Staubli VAL3: stop.pgx

program stop()
// Stop motion and preserve suction
begin
  resetMotion()
  blowOn = false
  if physicalRun
    taskKill("physicalIO")
    io:bOut1 = false
  endIf
  // Preserve suction so a held part is not released by STOP.
  cycleStep = -1
  putln("Stopped - empty the destinations before restarting")
end
